// TIA Portal V20 export
// export: Created 2026-10-12T15:48:32.5728389Z, ExportSetting WithDefaults, DisplayName Totally Integrated Automation Portal, DisplayVersion V20, DisplayName TIA Portal Openness, DisplayVersion V20, DisplayName TIA Portal Teamcenter Gateway, DisplayVersion V20, DisplayName TIA Portal Version Control Interface, DisplayVersion V20, DisplayName SINAMICS Startdrive Advanced, DisplayVersion V20 SP1 Update 2, DisplayName SINAMICS Startdrive G110M, G120, G120C, G120D, G120P, G115D, DisplayVersion V20 SP1 Update 2, DisplayName SINAMICS Startdrive G130, G150, S120, S150, SINAMICS MV, G220, S200, S210, DisplayVersion V20 SP1 Update 2, DisplayName STEP 7 Professional, DisplayVersion V20, DisplayName STEP 7 Safety, DisplayVersion V20, DisplayName WinCC Basic/Comfort/Advanced, DisplayVersion V20, DisplayName WinCC Professional, DisplayVersion V20, DisplayName WinCC Unified, DisplayVersion V20
FUNCTION "FRK_PartEvent" : Void   // FC71, SCL
{ S7_Optimized_Access := 'TRUE' }
VERSION : 0.1
// stored: AutoNumber true, IsIECCheckEnabled false, SetENOAutomatically false, UDAEnableTagReadback false
   VAR_INPUT
      Reason : DInt;
      Uid : String;
      SourcePath : String;
   END_VAR
   VAR_IN_OUT
      AlarmLog : "FRK_AlarmLog";
   END_VAR
   VAR_TEMP
      Description : WString[255];
   END_VAR
BEGIN

   CASE #Reason OF
       2024:
           #Description := WSTRING#'std.event.partReceived: ';
       2025:
           #Description := WSTRING#'std.event.partProcessingStarted: ';
       2026:
           #Description := WSTRING#'std.event.partProcessed: ';
       2027:
           #Description := WSTRING#'std.event.partAborted: ';
       ELSE
           #Description := WSTRING#'';
   END_CASE;
   #Description := CONCAT(IN1 := #Description, IN2 := STRING_TO_WSTRING(#Uid));
   "FRK_AlarmMessage"(AlarmLog := #AlarmLog,
                      Reason := #Reason,
                      Description := #Description,
                      SourcePath := STRING_TO_WSTRING(#SourcePath));
END_FUNCTION
